(* Sesnor Mismatch Detection *)

PROGRAM main
  VAR
    InputA AT %IX0.3 : BOOL;
    InputB AT %IX0.5 : BOOL;
    Output AT %MX0.3 : BOOL;
  END_VAR

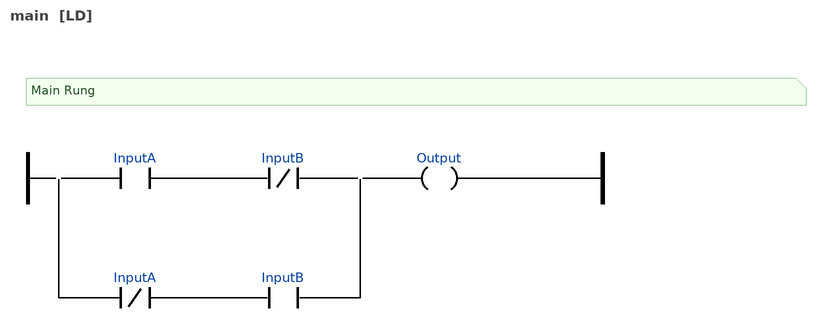
(* LD diagram, written out as Structured Text *)
(* Main Rung *)
Output := NOT InputA AND InputB OR InputA AND NOT InputB;
END_PROGRAM
